Staubli VAL3: IFedit.pgx

program IFedit(num x_nIndex)
begin
  call prog:editIF(sSelProg,x_nIndex,sIFType,sIFIndex,nIFValue,sANDOR1,sANDOR2,bToSave)
end
